// Motor 4 RETICLE VERT Y (SP1L0-KMONO-MMS-04)
//Main.M52.bLimitForwardEnable  := bM4CWLimit;    //(+Y)
//Main.M52.bLimitBackwardEnable := bM4CCWLimit;    //(-Y)
Main.M52.nEnableMode          := Enum_StageEnableMode.ALWAYS;
Main.M52.bHardwareEnable      := TRUE;
Main.M52.bPowerSelf           := TRUE;
fbMotion4(stMotionStage:=Main.M52);
//fbFFO4(stMotionStage := Main.M52,
//       fbFFHWO := GVL.fbFastFaultOutput1);
// Andy says: trip reticle if not OUT
// OUT is 1.55843, in is high limit switch
// NOTE: we don't have an encoder or an LVDT on this axis! We will use the out switch
bRetOut := NOT Main.M52.bLimitForwardEnable;
fbRetFFO(
    i_xOk := bRetOut,
    i_xAutoReset := TRUE,
    i_DevName := Main.M52.sName,
    i_Desc := 'Reticle not OUT (y>0)',
    io_fbFFHWO := GVL.fbFastFaultOutput1);

// Motor 5 DIODE HORIZ X (SP1L0-KMONO-MMS-05)
//Main.M53.bLimitForwardEnable  := bM5CCWLimit;    //(+X)
//Main.M53.bLimitBackwardEnable := bM5CWLimit;    //(-X)
Main.M53.nEnableMode          := Enum_StageEnableMode.DURING_MOTION;
Main.M53.bHardwareEnable      := TRUE;
Main.M53.bPowerSelf           := TRUE;
fbMotion5(stMotionStage:=Main.M53);

// Motor 6 DIODE VERT Y (SP1L0-KMONO-MMS-06)
//Main.M54.bLimitForwardEnable  := bM6CWLimit;    //(+Y)
//Main.M54.bLimitBackwardEnable := bM6CCWLimit;    //(-Y)
Main.M54.nEnableMode          := Enum_StageEnableMode.ALWAYS;
Main.M54.bHardwareEnable      := TRUE;
Main.M54.bPowerSelf           := TRUE;
fbMotion6(stMotionStage:=Main.M54);
//fbFFO6(stMotionStage := Main.M54,
//       fbFFHWO := GVL.fbFastFaultOutput1);
// Andy says trip if NOT IN or NOT OUT
// Andy says trip if IN AND NOT (7.7 to 8.9 keV)
// IN is 0, OUT is 98.5
bDiodeOut := Main.M54.stAxisStatus.fActPosition > 96.5;
bDiodeIn := Main.M54.stAxisStatus.fActPosition < 2;
fbDiodeFFOAtPos(
    i_xOk := bDiodeOut XOR bDiodeIn,
    i_xAutoReset := TRUE,
    i_DevName := Main.M54.sName,
    i_Desc := 'Diode between states.',
    io_fbFFHWO := GVL.fbFastFaultOutput1);
fbDiodeFFOEnergy(
    i_xOk := bEnergyOk OR NOT bDiodeIn,
    i_xReset := bDiodeOut OR (bDiodeIn AND bEnergyOk),
    i_xAutoReset := TRUE,
    i_DevName := Main.M54.sName,
    //i_Desc := 'Unsafe eV Range',
    i_Desc := 'Override if 7.7-8.9keV',
    io_fbFFHWO := GVL.fbFastFaultOutput1);

END_PROGRAM

// ---- POUs/PRG_3_PMPS_POST.TcPOU
PROGRAM PRG_3_PMPS_POST
VAR
    fbArbiterIO: FB_SubSysToArbiter_IO;
END_VAR

GVL.fbFastFaultOutput1.Execute();
GVL.fbFastFaultOutput2.Execute();

fbArbiterIO(
    Arbiter:=GVL.fbArbiter,
    fbFFHWO:=GVL.fbFastFaultOutput1);

END_PROGRAM

// ---- POUs/PRG_4_LOG.TcPOU
PROGRAM PRG_4_LOG
VAR
    fbLogHandler: FB_LogHandler;
END_VAR

fbLogHandler();

END_PROGRAM

// ---- Temp/FB_MPA.TcPOU
FUNCTION_BLOCK FB_MPA
VAR_INPUT
    (*EPS Interlock Bits*)
    ibInsertOK: BOOL;
    ibRetractOK: BOOL;
    ibPMPS_OK:BOOL;
    ibOverrideInterlock:BOOL; (*if true interlocks are ignored*)
    // Reset fault
    {attribute 'pytmc' := '
    pv: FF_Reset
    '}
    i_xReset: BOOL;
    sName: STRING;
    bEnableFF: BOOL := TRUE;
END_VAR
VAR_OUTPUT
    {attribute 'pytmc' := '
    pv:
    '}
    q_stAct     :    ST_MPA;
    {attribute 'pytmc' := '
    pv: MPS_FAULT
    '}
    xMPS_OK:BOOL;
    {attribute 'pytmc' := '
    pv: MOT_DONE
    '}
    xDone:Bool; // Motion is Done
END_VAR
VAR_IN_OUT
    io_fbFFHWO    :    FB_HardwareFFOutput;
END_VAR
VAR
    // PMPS
    fbFF    :    FB_FastFault :=(
        i_xAutoReset := TRUE,
        i_Desc := 'Device is moving',
        i_TypeCode := 16#1010);

    (*Init*)
    xFirstPass    :    BOOL;
    fbFSInit        :    R_TRIG;

    (* Timeouts*)
    tTimeOutDuration: TIME:= T#5S;
    tInserttimeout: TON;
    tRetracttimeout:TON;

    (*IO*)
    i_xInsertedLS    AT%I*: BOOL;
    i_xRetractedLS    AT%I*: BOOL;
    q_xInsert_DO    AT%Q*: BOOL;
    q_xRetract_DO    AT%Q*: BOOL;

    (* Reset Triggers *)
    rtInsert: R_TRIG;
    rtRemove: R_TRIG;
END_VAR


(*Initialize*)
fbFSInit( CLK := TRUE, Q => xFirstPass);
(*IO Mapping*)
ACT_IO();

IF xFirstPass THEN
    q_stAct.eState := INVALID;
    q_stAct.bRetract_SW := FALSE;
    q_stAct.bInsert_SW := FALSE;
END_IF


(* Manage States*)
IF q_stAct.i_bInLS AND  q_stAct.i_bOutLS THEN
    q_stAct.eState:=INVALID;
ELSIF NOT q_stAct.i_bInLS AND q_stAct.i_bOutLS THEN
    q_stAct.eState:=RETRACTED;
ELSIF q_stAct.i_bInLS AND NOT q_stAct.i_bOutLS THEN
    q_stAct.eState:=INSERTED;
ELSIF NOT q_stAct.i_bInLS AND NOT q_stAct.i_bOutLS THEN
    q_stAct.eState:=MOVING;
ELSE
    q_stAct.eState:=INVALID;
END_IF

(*Set the Done signal*)
xDone := (q_stAct.bRetract_SW AND q_stAct.eState=RETRACTED) OR (q_stAct.eState=INSERTED AND q_stAct.bInsert_SW);


(*MPS FAULT*)
(**)
xMPS_OK := (q_stAct.bRetract_SW AND i_xRetractedLS) XOR (i_xInsertedLS AND q_stAct.bInsert_SW);
//xMPS_OK := i_xRetractedLS XOR i_xInsertedLS;
//xMPS_OK := (q_stAct.eState=RETRACTED) OR (q_stAct.eState=INSERTED);
//xMPS_OK := (q_stAct.eState=RETRACTED) ;

(*PMPS PERMISSION*)

(* Reset the other command bit when one goes high *)
rtInsert(CLK:=q_stAct.bInsert_SW);
IF rtInsert.Q THEN
    q_stAct.bRetract_SW := FALSE;
END_IF
rtRemove(CLK:=q_stAct.bRetract_SW);
IF rtRemove.Q THEN
    q_stAct.bInsert_SW := FALSE;
END_IF

(* Can't have bRetract_SW and  bInsert_SW both be true*)
If (q_stAct.bRetract_SW) and (q_stAct.bInsert_SW) THEN
    q_stAct.bRetract_SW := FALSE;
    q_stAct.bInsert_SW := FALSE;
END_IF

(* Make the state consistent if we can *)
IF NOT (q_stAct.bRetract_SW OR q_stAct.bInsert_SW) THEN
    IF q_stAct.eState = RETRACTED THEN
        q_stAct.bRetract_SW := TRUE;
    ELSIF q_stAct.eState = INSERTED THEN
        q_stAct.bInsert_SW := TRUE;
    END_IF
END_IF

q_stAct.bRetractOK := ibRetractOK;
q_stAct.bInsertOK := ibInsertOK;

(*Actuate the device*)
q_stAct.q_bRetract := q_stAct.bRetractOK AND q_stAct.bRetract_SW;
q_stAct.q_bInsert := q_stAct.bInsertOK AND q_stAct.bInsert_SW;

IF q_stAct.q_bInsert THEN
    q_stAct.q_bRetract := FALSE;
    q_stAct.bRetract_SW:= FALSE;
ELSIF q_stAct.q_bRetract THEN
    q_stAct.q_bInsert := FALSE;
    q_stAct.bInsert_SW:= FALSE;
END_IF;




(*Timers*)
tInserttimeout(IN:= q_stAct.q_bInsert, PT := tTimeOutDuration );
tRetracttimeout(IN:= q_stAct.q_bRetract, PT := tTimeOutDuration);

///Check moving postion timout
IF NOT q_stAct.i_bInLS AND tInserttimeout.Q THEN
    q_stAct.bErrorPresent := TRUE;
ELSIF NOT q_stAct.i_bOutLS AND tRetracttimeout.Q THEN
    q_stAct.bErrorPresent := TRUE;
END_IF

(*FAST FAULT*)
IF bEnableFF THEN
    fbFF(i_DevName := sName,
        i_xOK := xMPS_OK,
        i_xReset := i_xReset,
        io_fbFFHWO := io_fbFFHWO);
END_IF

(*Soft IO Mapping*)
ACT_IO();

ACTION ACT_IO:
(*Inputs*)
q_stAct.i_bInLS :=  i_xInsertedLS;
q_stAct.i_bOutLS := i_xRetractedLS;

(*outputs*)
q_xInsert_DO:=q_stAct.q_bInsert;
q_xRetract_DO:=q_stAct.q_bRetract;
END_ACTION

END_FUNCTION_BLOCK

// ---- Temp/FB_BasicAxisFFO.TcPOU
FUNCTION_BLOCK FB_BasicAxisFFO
(*
    Placeholder FFO logic for no beam allowed, pre-comissioning

    Fast fault is applied if the axis is moving.
*)
VAR_IN_OUT
    Axis: AXIS_REF;
    fbFFHWO: FB_HardwareFFOutput;
END_VAR
VAR_INPUT
    sName: STRING;
END_VAR
VAR_OUTPUT
    bIsNotMoving: BOOL;
END_VAR
VAR
    fbFF: FB_FastFault := (i_Desc := 'Device is moving',
                           i_TypeCode := 16#2100,
                           i_xAutoReset := TRUE);
END_VAR

bIsNotMoving := NOT Axis.Status.Moving;
fbFF(i_DevName := sName,
     i_xOK := bIsNotMoving,
     io_fbFFHWO := fbFFHWO);

END_FUNCTION_BLOCK

// ---- Temp/FB_BasicMotionStageAltFFO.TcPOU
FUNCTION_BLOCK FB_BasicMotionStageAltFFO
(*
    Alternative to FB_BasicMotionStageFFO for an arbitrary out condition

    Sometimes the out limits is not what we want to use for proto-mps
*)
VAR_IN_OUT
    stMotionStage: DUT_MotionStage;
    fbFFHWO: FB_HardwareFFOutput;
END_VAR
VAR_INPUT
    sName: STRING;
    bFFOk: BOOL;
END_VAR
VAR_OUTPUT
    bIsOut: BOOL;
    bIsNotMoving: BOOL;
END_VAR
VAR
    fbBasicAxisFFO: FB_BasicAxisFFO := (sName := sName);
    fbFF: FB_FastFault := (i_Desc := 'Device is not out',
                           i_TypeCode := 16#2200,
                           i_xAutoReset := TRUE);
END_VAR

fbBasicAxisFFO(Axis := stMotionStage.Axis,
               fbFFHWO := fbFFHWO,
               sName := sName,
               bIsNotMoving => bIsNotMoving);

fbFF(i_DevName := sName,
     i_xOK := bFFOk,
     io_fbFFHWO := fbFFHWO);

END_FUNCTION_BLOCK

// ---- Temp/FB_BasicMotionStageFFO.TcPOU
FUNCTION_BLOCK FB_BasicMotionStageFFO
(*
    Placeholder FFO logic for no beam allowed, pre-comissioning

    Fast fault is applied if the motor is moving or is not at the out switch.
*)
VAR_IN_OUT
    stMotionStage: DUT_MotionStage;
    fbFFHWO: FB_HardwareFFOutput;
END_VAR
VAR_INPUT
    sName: STRING;
    bForwardIsOut: BOOL := TRUE;
END_VAR
VAR_OUTPUT
    bIsOut: BOOL;
    bIsNotMoving: BOOL;
END_VAR
VAR
    fbBasicAxisFFO: FB_BasicAxisFFO := (sName := sName);
    fbFF: FB_FastFault := (i_Desc := 'Device is not out',
                           i_TypeCode := 16#2200,
                           i_xAutoReset := TRUE);
END_VAR

fbBasicAxisFFO(Axis := stMotionStage.Axis,
               fbFFHWO := fbFFHWO,
               sName := sName,
               bIsNotMoving => bIsNotMoving);

IF bForwardIsOut THEN
    bIsOut := NOT stMotionStage.bLimitForwardEnable;
ELSE
    bIsOut := NOT stMotionStage.bLimitBackwardEnable;
END_IF

fbFF(i_DevName := sName,
     i_xOK := bIsOut,
     io_fbFFHWO := fbFFHWO);

END_FUNCTION_BLOCK

// ---- Temp/FB_DoubleActingMPA.TcPOU
FUNCTION_BLOCK FB_DoubleActingMPA
VAR_IN_OUT
    iq_MPA : DUT_DoubleActPneumaticActuator;
END_VAR

VAR


END_VAR


///Check valve postion



IF iq_MPA.i_xInsertLS AND iq_MPA.i_xRetractLS THEN
    iq_MPA.eState:=INVALID;
ELSIF NOT iq_MPA.i_xInsertLS AND iq_MPA.i_xRetractLS AND iq_MPA.q_xRetractDO THEN
    iq_MPA.eState:=RETRACTED;
ELSIF iq_MPA.i_xInsertLS AND NOT iq_MPA.i_xRetractLS AND NOT iq_MPA.q_xInsertDO THEN
    iq_MPA.eState:=INSERTED;
ELSIF NOT iq_MPA.i_xInsertLS AND NOT iq_MPA.i_xInsertLS THEN
    iq_MPA.eState:=MOVING;
ELSE
    iq_MPA.eState:=INVALID;
END_IF



IF iq_MPA._xInsertSW  THEN
    iq_MPA._xRetractSW := FALSE;
    iq_MPA.q_xRetractDO := FALSE;
    iq_MPA.q_xInsertDO := TRUE;
END_IF

IF iq_MPA._xRetractSW THEN
    iq_MPA._xInsertSW := FALSE;
    iq_MPA.q_xInsertDO:= FALSE;
    iq_MPA.q_xRetractDO := TRUE;
END_IF

END_FUNCTION_BLOCK

// ---- Temp/FB_SimMotor.TcPOU
FUNCTION_BLOCK FB_SimMotor
VAR_IN_OUT
    stMotionStage: DUT_MotionStage;
END_VAR
VAR
    fbMotionStage: FB_MotionStage;
END_VAR

stMotionStage.bLimitBackwardEnable := TRUE;
stMotionStage.bLimitForwardEnable := TRUE;
stMotionStage.bHardwareEnable := TRUE;
stMotionStage.bPowerSelf := TRUE;
stMotionStage.nEnableMode := ENUM_StageEnableMode.ALWAYS;
fbMotionStage(stMotionStage := stMotionStage);

END_FUNCTION_BLOCK

// ---- Temp/FB_SLITS_POWER_1.TcPOU
FUNCTION_BLOCK FB_SLITS_POWER_1
VAR_IN_OUT
    stTopBlade: DUT_MotionStage;
    stBottomBlade: DUT_MotionStage;
    stNorthBlade: DUT_MotionStage;
    stSouthBlade: DUT_MotionStage;
END_VAR
VAR_INPUT
    fPosTopBlade: LREAL;
    fPosBottomBlade: LREAL;
    fPosNorthBlade: LREAL;
    fPosSouthBlade: LREAL;
    bExecuteMotion:bool ;
END_VAR
VAR_OUTPUT
END_VAR
VAR
    fbTopBlade: FB_MotionStage;
    fbBottomBlade: FB_MotionStage;
    fbNorthBlade: FB_MotionStage;
    fbSouthBlade: FB_MotionStage;

    {attribute 'pytmc' := '
        pv: FSW
    '}
    fbFlowSwitch: FB_XTES_Flowswitch;


    //RTDs
    {attribute 'pytmc' := '
        pv: TOP:RTD:01
    '}
    RTD_TOP_1: FB_ThermoCouple;
    {attribute 'pytmc' := '
        pv: TOP:RTD:02
    '}
    RTD_TOP_2: FB_ThermoCouple;
    {attribute 'pytmc' := '
        pv: BOTTOM:RTD:01
    '}
    RTD_Bottom_1: FB_ThermoCouple;
    {attribute 'pytmc' := '
        pv: BOTTOM:RTD:02
    '}
    RTD_Bottom_2: FB_ThermoCouple;

    {attribute 'pytmc' := '
        pv: NORTH:RTD:01
    '}
    RTD_North_1: FB_ThermoCouple;
    {attribute 'pytmc' := '
        pv: NORTH:RTD:02
    '}
    RTD_North_2: FB_ThermoCouple;
    {attribute 'pytmc' := '
        pv: SOUTH:RTD:01
    '}
    RTD_South_1: FB_ThermoCouple;
    {attribute 'pytmc' := '
        pv: SOUTH:RTD:02
    '}
    RTD_South_2: FB_ThermoCouple;

    fSmallDelta: LREAL := 0.01;
    fBigDelta: LREAL := 10;
    fMaxVelocity: LREAL := 0.33;
    fHighAccel: LREAL := 0.8;
    fLowAccel: LREAL := 0.1;

    stTop: DUT_PositionState;
    stBOTTOM: DUT_PositionState;
    stNorth: DUT_PositionState;
    stSouth: DUT_PositionState;

    {attribute 'pytmc' := 'pv: TOP'}
    fbTop: FB_StatePTPMove;
    {attribute 'pytmc' := 'pv: BOTTOM'}
    fbBottom: FB_StatePTPMove;
    {attribute 'pytmc' := 'pv: NORTH'}
    fbNorth: FB_StatePTPMove;
    {attribute 'pytmc' := 'pv: SOUTH'}
    fbSouth: FB_StatePTPMove;


END_VAR

// Instantiate Function block for all the blades
fbTopBlade(stMotionStage:=stTopBlade);
fbBottomBlade(stMotionStage:=stBottomBlade);
fbNorthBlade(stMotionStage:=stNorthBlade);
fbSouthBlade(stMotionStage:=stSouthBlade);

//  no STO
stTopBlade.bHardwareEnable := TRUE;
stBottomBlade.bHardwareEnable := TRUE;
stNorthBlade.bHardwareEnable := TRUE;
stSouthBlade.bHardwareEnable := TRUE;
stTopBlade.bPowerSelf :=TRUE;
stBottomBlade.bPowerSelf :=TRUE;
stNorthBlade.bPowerSelf :=TRUE;
stSouthBlade.bPowerSelf :=TRUE;

//RTDs
RTD_TOP_1();
RTD_TOP_2();
RTD_Bottom_1();
RTD_Bottom_2();
RTD_North_1();
RTD_North_2();
RTD_South_1();
RTD_South_2();

//Flow Switch
fbFlowSwitch();


// PTP Motion for each blade

stTop.sName := 'Top';
stTop.fPosition := fPosTopBlade;
stTop.fDelta := fSmallDelta;
stTop.fVelocity := fMaxVelocity;
stTop.fAccel := fHighAccel;
stTop.fDecel := fHighAccel;

stBOTTOM.sName := 'Bottom';
stBOTTOM.fPosition := fPosBottomBlade;
stBOTTOM.fDelta := fSmallDelta;
stBOTTOM.fVelocity := fMaxVelocity;
stBOTTOM.fAccel := fHighAccel;
stBOTTOM.fDecel := fHighAccel;

stNorth.sName := 'North';
stNorth.fPosition := fPosNorthBlade;
stNorth.fDelta := fSmallDelta;
stNorth.fVelocity := fMaxVelocity;
stNorth.fAccel := fHighAccel;
stNorth.fDecel := fHighAccel;

stSouth.sName := 'South';
stSouth.fPosition := fPosSouthBlade;
stSouth.fDelta := fSmallDelta;
stSouth.fVelocity := fMaxVelocity;
stSouth.fAccel := fHighAccel;
stSouth.fDecel := fHighAccel;

//fbTop.bExecute := fbBottom.bExecute :=fbNorth.bExecute := fbSouth.bExecute := bExecuteMotion;

fbTop(
    stPositionState:=stTop,
    bMoveOk:=TRUE,
    stMotionStage:=stTopBlade);

fbBottom(
    stPositionState:=stBOTTOM,
    bMoveOk:=TRUE,
    stMotionStage:=stBottomBlade);

fbNorth(
    stPositionState:=stNorth,
    bMoveOk:=TRUE,
    stMotionStage:=stNorthBlade);

fbSouth(
    stPositionState:=stSouth,
    bMoveOk:=TRUE,
    stMotionStage:=stSouthBlade);

END_FUNCTION_BLOCK
